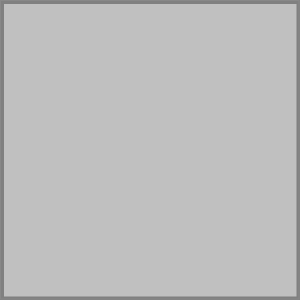
VISUALIZATION viz_HMI_Piston  // 300x300
VAR_INPUT
	bLock_HMI: BOOL;
END_VAR
    Rectangle (0,0 300x300), invisible if: TRUE
END_VISUALIZATION

(* stored: Version 1.1.0.1, ProductVersion 3.1.4024.13
   Visu viz_HMI_Piston: Id {fa1b94a3-45a7-4c31-8230-f8d8dacbd140} *)
